// Ein Niederhalter (DFM-50, monostabiles 5/2-Ventil, Grundstellung OFFEN, Sensor nur auf Endlage OFFEN).
// „Geklemmt“ = Endlage OFFEN verlassen, Druck in Ordnung und Schaltzeit abgelaufen [Langfeld].
FUNCTION_BLOCK FB_Clamp
VAR_INPUT
    bSensorOpen : BOOL;
    bPressureOk : BOOL;
    bForceOpen : BOOL;      // Not-Halt: Ventil aus (Pneumatik wird ohnehin entlüftet)
END_VAR
VAR_OUTPUT
    bValve : BOOL;
    eState : E_ClampState := E_ClampState.Unknown;
    bTimeoutFault : BOOL;
    bPressureFault : BOOL;
    fLastSwitchTime_ms : LREAL;
END_VAR
VAR
    bCmdClose : BOOL;
    tonSwitch : TON;
    tonTimeout : TON;
    tStart : TIME;
END_VAR

IF bForceOpen THEN
    bCmdClose := FALSE;
END_IF
bValve := bCmdClose;
tonSwitch(IN := bCmdClose, PT := GVL_Config.tClampSwitch);
tonTimeout(IN := (eState = E_ClampState.Closing) OR (eState = E_ClampState.Opening), PT := GVL_Config.tClampTimeout);

CASE eState OF
E_ClampState.Unknown:
    IF bCmdClose THEN
        eState := E_ClampState.Closing;
    ELSIF bSensorOpen THEN
        eState := E_ClampState.Open;
    ELSE
        eState := E_ClampState.Opening;
    END_IF

E_ClampState.Open:
    IF bCmdClose THEN
        eState := E_ClampState.Closing;
        tStart := TIME();
    ELSIF NOT bSensorOpen THEN
        eState := E_ClampState.Opening;     // Endlage verloren: neu überwachen
    END_IF

E_ClampState.Closing:
    IF NOT bCmdClose THEN
        eState := E_ClampState.Opening;
        tStart := TIME();
    ELSIF tonSwitch.Q AND NOT bSensorOpen AND bPressureOk THEN
        eState := E_ClampState.Clamped;
        fLastSwitchTime_ms := TIME_TO_LREAL(TIME() - tStart);
    ELSIF tonTimeout.Q THEN
        eState := E_ClampState.Fault;
        bTimeoutFault := TRUE;
    END_IF

E_ClampState.Clamped:
    IF NOT bCmdClose THEN
        eState := E_ClampState.Opening;
        tStart := TIME();
    ELSIF NOT bPressureOk THEN
        eState := E_ClampState.Fault;
        bPressureFault := TRUE;
    END_IF

E_ClampState.Opening:
    IF bCmdClose THEN
        eState := E_ClampState.Closing;
        tStart := TIME();
    ELSIF bSensorOpen THEN
        eState := E_ClampState.Open;
        fLastSwitchTime_ms := TIME_TO_LREAL(TIME() - tStart);
    ELSIF tonTimeout.Q THEN
        eState := E_ClampState.Fault;
        bTimeoutFault := TRUE;
    END_IF

E_ClampState.Fault:
    // bleibt bis ResetFault(); Ventil folgt weiter dem Kommando
    ;
END_CASE

METHOD Close : BOOL
VAR_INPUT
END_VAR
bCmdClose := TRUE;
Close := TRUE;
END_METHOD

METHOD Open : BOOL
VAR_INPUT
END_VAR
bCmdClose := FALSE;
Open := TRUE;
END_METHOD

METHOD ResetFault : BOOL
VAR_INPUT
END_VAR
IF eState = E_ClampState.Fault THEN
    bTimeoutFault := FALSE;
    bPressureFault := FALSE;
    eState := E_ClampState.Unknown;
END_IF
ResetFault := TRUE;
END_METHOD

METHOD IsOpen : BOOL
VAR_INPUT
END_VAR
IsOpen := eState = E_ClampState.Open;
END_METHOD

METHOD IsClamped : BOOL
VAR_INPUT
END_VAR
IsClamped := eState = E_ClampState.Clamped;
END_METHOD

METHOD IsCommandedClosed : BOOL
VAR_INPUT
END_VAR
IsCommandedClosed := bCmdClose;
END_METHOD

END_FUNCTION_BLOCK

(* stored: Version 1.1.0.1
   POU FB_Clamp: Id {936507bc-9160-5df3-aa91-1edf155c1c67}, SpecialFunc None
   Method Close: Id {aad6d455-139d-5ea1-8369-9a92d496da9e}
   Method Open: Id {21611771-ffff-5d6a-a327-7035c70542d6}
   Method ResetFault: Id {6567cef7-68e8-5e23-9015-53211eb22c47}
   Method IsOpen: Id {c192c712-86b8-56a1-8001-788434a7db8a}
   Method IsClamped: Id {055e9054-64db-583f-80e9-f341b7a63307}
   Method IsCommandedClosed: Id {cd878e4e-b457-5eba-b170-b1b46d63c8ae} *)
